Yaskawa INFORM job: CALIBVISION.JBI

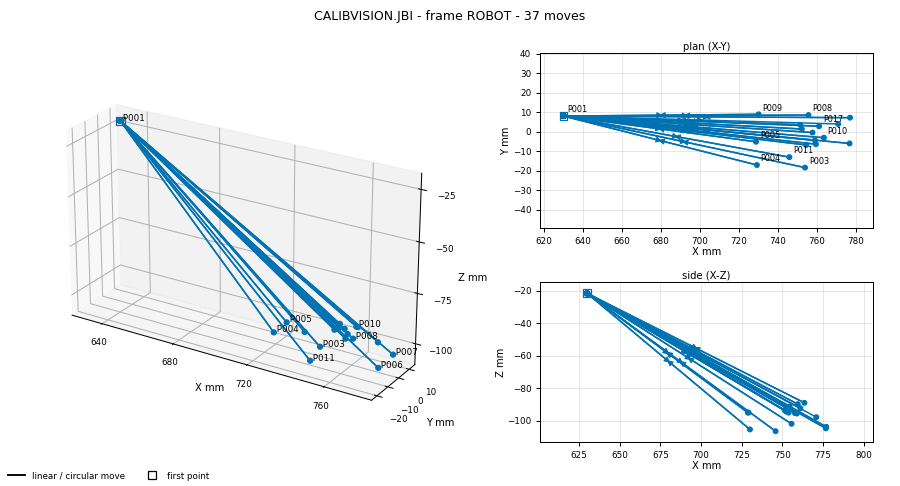
[picture p0: tool path of CALIBVISION.JBI in frame ROBOT, 37 of 38 moves have a stored position in this frame; points joined in program order, loops and branches not executed]
/JOB
//NAME CALIBVISION
///FOLDERNAME FOLDER003
//POS
///NPOS 1,0,0,19,0,0
///TOOL 1
///POSTYPE PULSE
///PULSE
C00000=-7868,-19030,-10844,-11154,-67763,7913
///POSTYPE ROBOT
///RECTAN
///RCONF 0,0,0,0,0,0,0,0,0,0,0,0,0,0,0,0,0,0,0,0,0,0,0,0
P00001=629.883,8.042,-21.694,-154.9112,52.6025,29.7528
P00002=629.627,8.031,-21.395,-154.9194,52.6073,29.7435
P00003=753.895,-18.403,-95.100,179.0147,0.9881,-3.6266
P00004=729.189,-17.091,-95.012,179.5704,3.1491,-3.5911
P00005=728.757,-5.152,-95.055,179.5608,3.1535,-3.5736
P00006=776.762,-6.009,-104.764,-174.3345,-0.2294,-3.5144
P00007=777.008,7.220,-103.781,-178.0279,-4.4731,-2.4061
P00008=755.683,8.551,-101.944,179.1931,-0.6151,-3.5050
P00009=730.061,8.946,-105.416,-176.1634,4.1381,-4.6170
P00010=763.595,-3.084,-89.028,166.6757,11.1463,-4.9576
P00011=745.860,-13.056,-106.500,-158.3053,3.8563,-0.2463
P00012=757.745,-0.414,-95.337,-179.5172,24.2328,-2.1533
P00013=759.483,-6.389,-89.840,172.3389,-15.9039,-2.7723
P00014=758.946,-4.455,-95.629,175.1183,-2.0647,-15.9599
P00015=754.520,-6.809,-91.368,175.1177,-2.0668,14.8104
P00016=751.436,3.569,-93.547,175.1246,-2.0642,-21.6342
P00017=761.103,2.831,-92.360,177.0136,-2.5401,7.3666
P00018=752.261,1.393,-94.364,-178.1918,0.5648,17.2122
P00019=770.910,3.984,-97.871,175.1225,-2.0691,24.6146
//INST
///DATE 2025/04/28 09:17
///ATTR SC,RW
///GROUP1 RB1
NOP
MOVL P001 V=20.0 PL=0
CALL JOB:CALIBPOSON
MOVL P001 V=5.0
MOVL P002 V=5.0 PL=0
CALL JOB:CALIBPOSON
MOVL P001 V=5.0
MOVL P003 V=5.0 PL=0
CALL JOB:CALIBPOSON
MOVL P001 V=5.0
MOVL P004 V=5.0 PL=0
CALL JOB:CALIBPOSON
MOVL P001 V=5.0
MOVL P005 V=5.0 PL=0
CALL JOB:CALIBPOSON
MOVL P001 V=5.0
MOVL P006 V=5.0 PL=0
CALL JOB:CALIBPOSON
MOVL P001 V=5.0
MOVL P007 V=5.0 PL=0
CALL JOB:CALIBPOSON
MOVL P001 V=5.0
MOVL P008 V=5.0 PL=0
CALL JOB:CALIBPOSON
MOVL P001 V=5.0
MOVL P009 V=5.0 PL=0
CALL JOB:CALIBPOSON
MOVL P001 V=5.0
MOVL P010 V=3.0 PL=0
CALL JOB:CALIBPOSON
MOVL P001 V=5.0
MOVL P011 V=3.0 PL=0
CALL JOB:CALIBPOSON
MOVL P001 V=5.0
MOVL P012 V=3.0 PL=0
CALL JOB:CALIBPOSON
MOVL P001 V=5.0
MOVL P013 V=3.0 PL=0
CALL JOB:CALIBPOSON
MOVL P001 V=5.0
MOVL P014 V=3.0 PL=0
CALL JOB:CALIBPOSON
MOVL P001 V=5.0
MOVL P015 V=3.0 PL=0
CALL JOB:CALIBPOSON
MOVL P001 V=5.0
MOVL P016 V=5.0 PL=0
CALL JOB:CALIBPOSON
MOVL P001 V=5.0
MOVL P017 V=5.0 PL=0
CALL JOB:CALIBPOSON
MOVL P001 V=5.0
MOVL P018 V=5.0 PL=0
CALL JOB:CALIBPOSON
MOVL P001 V=5.0
MOVL P019 V=5.0 PL=0
CALL JOB:CALIBPOSON
MOVL C00000
END
